(* IEC 61131-3 sources: BODAS-RC27-18_40/st/bodas_rc18_12_27_18_40/plc_logic/application/easyconfig_import/bds_in_legacy_ec, 7 files *)

(* ---- bds_in_aiv_signal_te-bds_in_aiv_signal_te.st ---- *)
(* --- Interface --- *)
{attribute 'qualified_only' := ''}
{attribute 'strict' := ''}
TYPE bds_in_aiv_signal_te :
(
	IN_AIV_START_SIGNALS := 16#500,
	IN_AIV_START := 16#4FF,
	K52,
	K60,
	K43,
	K54,
	K55,
	K37,
	K61,
	A21,
	A36,
	A37,
	A38,
	A39,
	K32,
	K30,
	K78,
	K76,
	K74,
	K77,
	K10,
	K75,
	K31,
	K34,
	A13,
	A40,
	A41,
	A42,
	A25,
	A26,
	A27,
	A14,
	A57,
	A28,
	A29,
	K11,
	K35,
	IN_AIV_NUM_SIGNALS,
	IN_AIV_FLEXIN_NUM_SIGNALS := K78
) UINT;
END_TYPE

(* ---- bds_in_di_signal_te-bds_in_di_signal_te.st ---- *)
(* --- Interface --- *)
{attribute 'qualified_only' := ''}
{attribute 'strict' := ''}
TYPE bds_in_di_signal_te :
(
	IN_DI_START_SIGNALS := 16#400,
	IN_DI_START := 16#3FF,
	K39,
	K38,
	K40,
	K41,
	K42,
	A43,
	K21,
	K22,
	IN_DI_NUM_SIGNALS
) UINT;
END_TYPE

(* ---- bds_in_fi_signal_te-bds_in_fi_signal_te.st ---- *)
(* --- Interface --- *)
{attribute 'qualified_only' := ''}
{attribute 'strict' := ''}
TYPE bds_in_fi_signal_te :
(
	IN_FI_START_SIGNALS := 16#700,
	IN_FI_START := 16#6FF,
	K39_VI,
	K38_VI,
	K40_VI,
	K41_VI,
	K42_VI,
	K45_VI,
	K44_VI,
	K65_VI,
	K63_VI,
	K64_VI,
	A36_VI,
	A37_VI,
	A38_VI,
	A39_VI,
	K55_VI,
	K61_VI,
	K30_VI,
	A43_VI,
	K53,
	K57,
	K58,
	K36,
	A22,
	A23,
	A24,
	IN_FI_NUM_SIGNALS,
	IN_FI_DSM_NUM_SIGNALS := K53
) UINT;
END_TYPE

(* ---- bds_in_phase_signal_te-bds_in_phase_signal_te.st ---- *)
(* --- Interface --- *)
{attribute 'qualified_only' := ''}
{attribute 'strict' := ''}
TYPE bds_in_phase_signal_te :
(
	IN_PHASE_START_SIGNALS := 16#900,
	IN_PHASE_START := 16#8FF,
	K54_VI_K37_VI,
	IN_PHASE_NUM_SIGNALS
) UINT;
END_TYPE

(* ---- bds_in_ri_signal_te-bds_in_ri_signal_te.st ---- *)
(* --- Interface --- *)
{attribute 'qualified_only' := ''}
{attribute 'strict' := ''}
TYPE bds_in_ri_signal_te :
(
	IN_RI_START_SIGNALS := 16#600,
	IN_RI_START := 16#5FF,
	K45,
	K44,
	K65,
	K63,
	K64,
	K33,
	IN_RI_NUM_SIGNALS
) UINT;
END_TYPE

(* ---- bds_in_sent_signal_te-bds_in_sent_signal_te.st ---- *)
(* --- Interface --- *)
{attribute 'qualified_only' := ''}
{attribute 'strict' := ''}
TYPE bds_in_sent_signal_te :
(
	IN_SENT_START_SIGNALS := 16#800,
	IN_SENT_START := 16#7FF,
	K59,
	K56,
	IN_SENT_NUM_SIGNALS
) UINT;
END_TYPE

(* ---- bds_in_legacy_ec_gvl-bds_in_legacy_ec_gvl.st ---- *)
(* --- Interface --- *)
{attribute 'qualified_only' := ''}
VAR_GLOBAL CONSTANT
	ACTIVATE_SHUNT_AIC_K39: UDINT := 0;
	ACTIVATE_SHUNT_AIC_K38: UDINT := 0;
	ACTIVATE_SHUNT_AIC_K40: UDINT := 0;
	ACTIVATE_SHUNT_AIC_K41: UDINT := 0;
	ACTIVATE_SHUNT_AIC_K42: UDINT := 0;
	ACTIVATE_SHUNT_AIC_K45: UDINT := 0;
	ACTIVATE_SHUNT_AIC_K44: UDINT := 0;
	ACTIVATE_SHUNT_AIC_K65: UDINT := 0;
	ACTIVATE_SHUNT_AIC_K63: UDINT := 0;
	ACTIVATE_SHUNT_AIC_K64: UDINT := 0;
	ACTIVATE_SHUNT_AIC_A36: UDINT := 0;
	ACTIVATE_SHUNT_AIC_A37: UDINT := 1;
	ACTIVATE_SHUNT_AIC_A38: UDINT := 0;
	ACTIVATE_SHUNT_AIC_A39: UDINT := 0;
	ACTIVATE_SHUNT1: UDINT := 0;
	ACTIVATE_SHUNT2: UDINT := 1;
	ACTIVATE_SHUNT3: UDINT := 0;
	ACTIVATE_SHUNT4: UDINT := 0;
	ACTIVATE_SHUNT5: UDINT := 1;
	ACTIVATE_SHUNT6: UDINT := 0;
	BDS_IN_AIV_32V_NUM_SIGNALS_D: UINT := bds_in_aiv_signal_te.A14;
	BDS_IN_FI_AIC_NUM_SIGNALS_D: UINT := bds_in_fi_signal_te.K55_VI;
END_VAR
